FUNCTION_BLOCK SENSOR_VOTER (* Migrated from IEC 61131-3 ST *)
  (* Standard: 61499-2 *)
  (* Version 1.0, 2026-11-06, st2fb *)
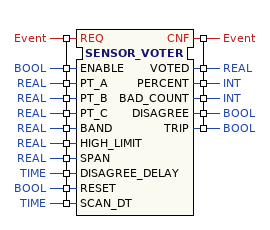
  EVENT_INPUT
    REQ WITH ENABLE, PT_A, PT_B, PT_C, BAND, HIGH_LIMIT, SPAN, DISAGREE_DELAY, RESET, SCAN_DT;
  END_EVENT
  EVENT_OUTPUT
    CNF WITH VOTED, PERCENT, BAD_COUNT, DISAGREE, TRIP;
  END_EVENT
  VAR_INPUT
    ENABLE : BOOL;
    PT_A : REAL;
    PT_B : REAL;
    PT_C : REAL;
    BAND : REAL;
    HIGH_LIMIT : REAL;
    SPAN : REAL;
    DISAGREE_DELAY : TIME;
    RESET : BOOL;
    SCAN_DT : TIME;
  END_VAR
  VAR_OUTPUT
    VOTED : REAL;
    PERCENT : INT;
    BAD_COUNT : INT;
    DISAGREE : BOOL;
    TRIP : BOOL;
  END_VAR
  VAR
    MIDDLE : REAL;
    OVER_HIGH : BOOL;
    ST2FB_NOW : TIME := T#0s;
    DT_IN : BOOL;
    DT_PT : TIME;
    DT_Q : BOOL;
    DT_ET : TIME;
    DT_STATE : INT;
    DT_PREV_IN : BOOL;
    DT_START_TIME : TIME;
    TL_S : BOOL;
    TL_R1 : BOOL;
    TL_Q1 : BOOL;
  END_VAR
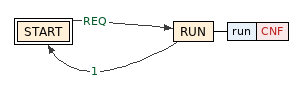
  EC_STATES
    START;
    RUN : run -> CNF;
  END_STATES
  EC_TRANSITIONS
    START TO RUN := REQ;
    RUN TO START := 1;
  END_TRANSITIONS
  ALGORITHM run IN ST:
ST2FB_NOW := ST2FB_NOW + SCAN_DT;
IF NOT ENABLE THEN
  DT_IN := FALSE;
  DT_PT := DISAGREE_DELAY;
  IF (DT_STATE = 0) AND NOT DT_PREV_IN AND DT_IN THEN
    DT_STATE := 1;
    DT_Q := FALSE;
    DT_START_TIME := ST2FB_NOW;
  ELSE
    IF NOT DT_IN THEN
      DT_ET := T#0s;
      DT_Q := FALSE;
      DT_STATE := 0;
    ELSIF DT_STATE = 1 THEN
      IF DT_START_TIME + DT_PT <= ST2FB_NOW THEN
        DT_STATE := 2;
        DT_Q := TRUE;
        DT_ET := DT_PT;
      ELSE
        DT_ET := ST2FB_NOW - DT_START_TIME;
      END_IF;
    END_IF;
  END_IF;
  DT_PREV_IN := DT_IN;
  DISAGREE := FALSE;
  BAD_COUNT := 0;
ELSE
  MIDDLE := MAX(MIN(PT_A, PT_B), MIN(MAX(PT_A, PT_B), PT_C));
  BAD_COUNT := 0;
  IF ABS(PT_A - MIDDLE) > BAND THEN
    BAD_COUNT := BAD_COUNT + 1;
  END_IF;
  IF ABS(PT_B - MIDDLE) > BAND THEN
    BAD_COUNT := BAD_COUNT + 1;
  END_IF;
  IF ABS(PT_C - MIDDLE) > BAND THEN
    BAD_COUNT := BAD_COUNT + 1;
  END_IF;

  DT_IN := BAD_COUNT > 0;
  DT_PT := DISAGREE_DELAY;
  IF (DT_STATE = 0) AND NOT DT_PREV_IN AND DT_IN THEN
    DT_STATE := 1;
    DT_Q := FALSE;
    DT_START_TIME := ST2FB_NOW;
  ELSE
    IF NOT DT_IN THEN
      DT_ET := T#0s;
      DT_Q := FALSE;
      DT_STATE := 0;
    ELSIF DT_STATE = 1 THEN
      IF DT_START_TIME + DT_PT <= ST2FB_NOW THEN
        DT_STATE := 2;
        DT_Q := TRUE;
        DT_ET := DT_PT;
      ELSE
        DT_ET := ST2FB_NOW - DT_START_TIME;
      END_IF;
    END_IF;
  END_IF;
  DT_PREV_IN := DT_IN;
  DISAGREE := DT_Q;

  VOTED := MIDDLE;
  PERCENT := REAL_TO_INT(100.0 * VOTED / SPAN);

  OVER_HIGH := (VOTED > HIGH_LIMIT) AND (BAD_COUNT < 2);
  TL_S := OVER_HIGH;
  TL_R1 := RESET;
  TL_Q1 := NOT TL_R1 AND (TL_S OR TL_Q1);
  TRIP := TL_Q1;
END_IF;
  END_ALGORITHM
END_FUNCTION_BLOCK
